PROGRAM main
  VAR
    run AT %QX0.1 : BOOL; (* Cell run permission, a self-holding output *)
    estop_active AT %QX0.2 : BOOL; (* E-stop loop is open right now *)
    reset_cmd AT %QX0.3 : BOOL; (* Reset accepted, only with the E-stop loop closed *)
    st_idle AT %QX0.4 : BOOL; (* State IDLE *)
    st_run AT %QX0.5 : BOOL; (* State RUN *)
    st_pick AT %QX0.6 : BOOL; (* State PICK *)
    st_place AT %QX0.7 : BOOL; (* State PLACE *)
    st_done AT %QX1.0 : BOOL; (* State DONE *)
    estop_latch AT %QX1.1 : BOOL; (* E-stop latched, cleared only by reset *)
    st_fault AT %QX1.2 : BOOL; (* State FAULT *)
    drive_alarm AT %QX1.3 : BOOL;
    start_pb AT %QX2.0 : BOOL; (* Start push button, 0.5 s pulse *)
    stop_pb AT %QX2.1 : BOOL; (* Stop push button, 0.5 s pulse *)
    estop_ok AT %QX2.2 : BOOL; (* E-stop loop healthy, 1 = closed *)
    reset_pb AT %QX2.3 : BOOL; (* Reset push button, 0.5 s pulse *)
    at_home AT %QX2.4 : BOOL; (* Arm is at the home pose *)
    cycle_done AT %QX2.5 : BOOL; (* All cubes sorted *)
    r_fault AT %QX2.6 : BOOL; (* Robot fault (IK failure or similar) *)
    ph_pick AT %QX2.7 : BOOL; (* Arm is in the pick phase *)
    ph_place AT %QX3.0 : BOOL; (* Arm is in the place phase *)
    arm_busy AT %QX3.1 : BOOL; (* Arm is moving (unused in the rungs) *)
    drive_fault AT %QX3.2 : BOOL;
    interrupted : BOOL; (* The arm left home under run and has not returned *)
    can_start : BOOL; (* Start interlock: at home or interrupted *)
  END_VAR

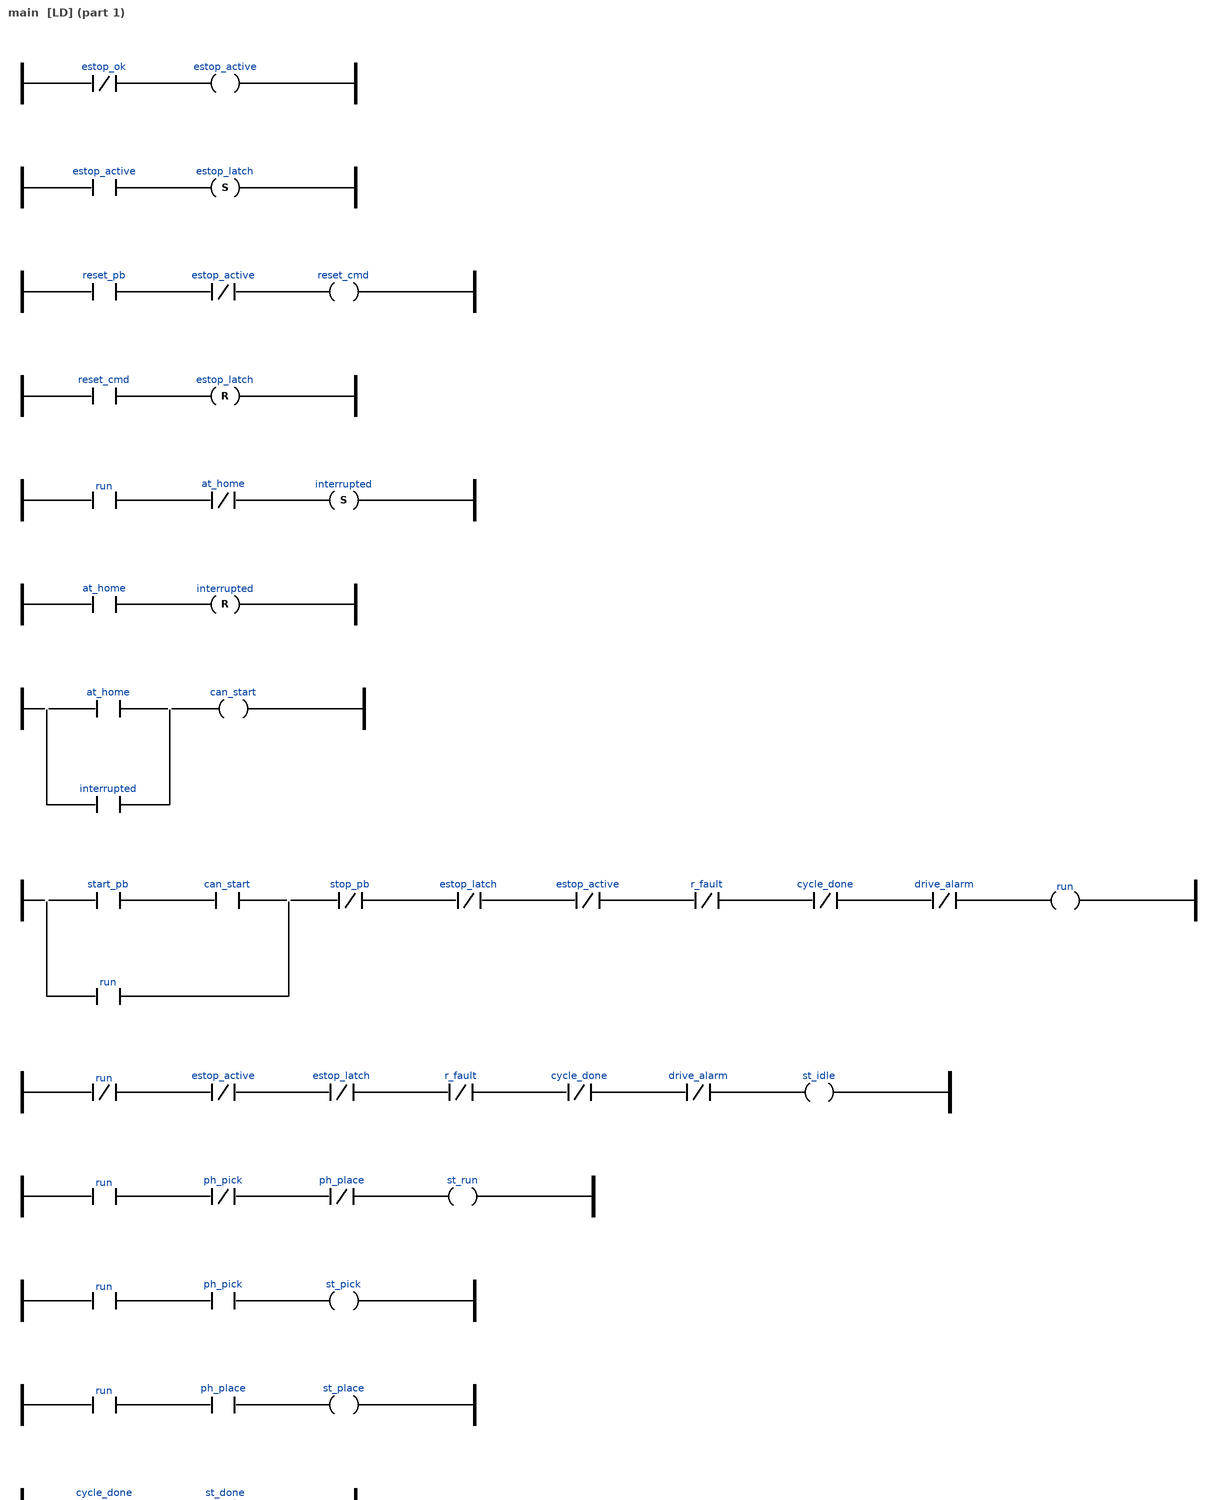
(* LD diagram, written out as Structured Text *)
estop_active := NOT estop_ok;
IF estop_active THEN estop_latch := TRUE; END_IF;
reset_cmd := reset_pb AND NOT estop_active;
IF reset_cmd THEN estop_latch := FALSE; END_IF;
IF run AND NOT at_home THEN interrupted := TRUE; END_IF;
IF at_home THEN interrupted := FALSE; END_IF;
can_start := at_home OR interrupted;
run := (run OR start_pb AND can_start) AND NOT stop_pb AND NOT estop_latch AND NOT estop_active AND NOT r_fault AND NOT cycle_done AND NOT drive_alarm;
st_idle := NOT run AND NOT estop_active AND NOT estop_latch AND NOT r_fault AND NOT cycle_done AND NOT drive_alarm;
st_run := run AND NOT ph_pick AND NOT ph_place;
st_pick := run AND ph_pick;
st_place := run AND ph_place;
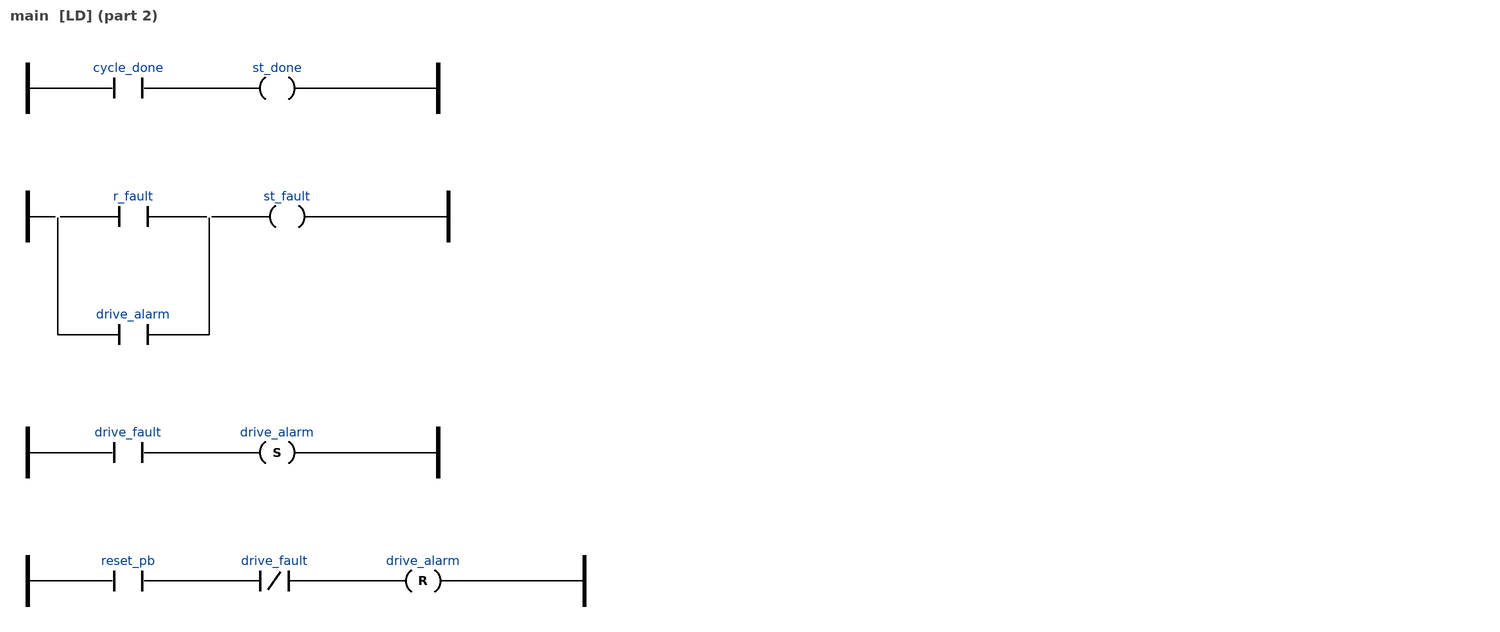
st_done := cycle_done;
st_fault := r_fault OR drive_alarm;
IF drive_fault THEN drive_alarm := TRUE; END_IF;
IF reset_pb AND NOT drive_fault THEN drive_alarm := FALSE; END_IF;
END_PROGRAM
